(* IEC 61131-3 sources: model-first-plc-agent-ai/results/T2-W-22, 2 files *)

(* ---- a1_code.st ---- *)
FUNCTION_BLOCK FillingRuntime
VAR_INPUT
    start : BOOL;
    stop : BOOL;
    LSH : BOOL;
    LSHH : BOOL;
    TimerDuration : TIME;
END_VAR
VAR_OUTPUT
    fill_valve : BOOL;
    discharge_valve : BOOL;
END_VAR
VAR
    x0 : BOOL := TRUE;
    x1 : BOOL := FALSE;
    timer_done : BOOL := FALSE;
    FillingTimer : TON;
END_VAR

(* Admit a start event only from the initial situation. *)
IF x0 AND start AND NOT stop AND NOT LSHH THEN
    x0 := FALSE;
    x1 := TRUE;
END_IF;

(* Timing begins in the same scan that x1 becomes active. *)
FillingTimer(IN := x1, PT := TimerDuration);
timer_done := FillingTimer.Q;

(* Terminate filling before updating the physical output commands. *)
IF x1 AND (stop OR LSHH OR timer_done) THEN
    x1 := FALSE;
    x0 := TRUE;

    (* Reset immediately so a subsequent start receives a fresh interval. *)
    FillingTimer(IN := FALSE, PT := TimerDuration);
    timer_done := FALSE;
END_IF;

fill_valve := x1;
discharge_valve := FALSE;

END_FUNCTION_BLOCK

PROGRAM Main
VAR
    StartCommand AT %IX100.0 : BOOL;
    StopCommand AT %IX100.1 : BOOL;
    LSH AT %IX100.2 : BOOL;
    LSHH AT %IX100.3 : BOOL;
    FillValve AT %QX100.0 : BOOL;
    DischargeValve AT %QX100.1 : BOOL;
END_VAR
VAR
    (* Configurable filling interval. *)
    TimerDuration : TIME := T#5s;
    StartEdge : R_TRIG;
    FillingControl : FillingRuntime;
END_VAR

StartEdge(CLK := StartCommand);

FillingControl(
    start := StartEdge.Q,
    stop := StopCommand,
    LSH := LSH,
    LSHH := LSHH,
    TimerDuration := TimerDuration
);

FillValve := FillingControl.fill_valve;
DischargeValve := FillingControl.discharge_valve;

END_PROGRAM

(* ---- a2_code.st ---- *)
FUNCTION_BLOCK FB_TimedTank
VAR_INPUT
    StartCommand : BOOL;
    StopCommand : BOOL;
    LSH : BOOL;
    LSHH : BOOL;
    TimerDuration : TIME;
END_VAR
VAR_OUTPUT
    fill_valve : BOOL;
    discharge_valve : BOOL;
END_VAR
VAR
    StartEdge : R_TRIG;
    FillingTimer : TON;
    CycleState : INT := 0;
    start : BOOL;
    stop : BOOL;
    timer_done : BOOL;
END_VAR

StartEdge(CLK := StartCommand);
start := StartEdge.Q;
stop := StopCommand;

IF stop THEN
    CycleState := 0;
ELSE
    CASE CycleState OF
        0:
            IF start AND NOT LSHH THEN
                CycleState := 1;
            END_IF;
        1:
            IF LSHH THEN
                CycleState := 0;
            END_IF;
    ELSE
        CycleState := 0;
    END_CASE;
END_IF;

(* Start timing in the same scan that the filling step becomes active. *)
FillingTimer(IN := (CycleState = 1), PT := TimerDuration);
timer_done := FillingTimer.Q;

IF (CycleState = 1) AND timer_done THEN
    CycleState := 0;

    (* Reset the owned timer immediately upon leaving the filling step. *)
    FillingTimer(IN := FALSE, PT := TimerDuration);
    timer_done := FillingTimer.Q;
END_IF;

fill_valve := (CycleState = 1);
discharge_valve := FALSE;

END_FUNCTION_BLOCK

PROGRAM Main
VAR
    StartCommand AT %IX100.0 : BOOL;
    StopCommand AT %IX100.1 : BOOL;
    LSH AT %IX100.2 : BOOL;
    LSHH AT %IX100.3 : BOOL;
    FillValve AT %QX100.0 : BOOL;
    DischargeValve AT %QX100.1 : BOOL;
END_VAR
VAR
    TankController : FB_TimedTank;
    TimerDuration : TIME := T#5s;
END_VAR

TankController(
    StartCommand := StartCommand,
    StopCommand := StopCommand,
    LSH := LSH,
    LSHH := LSHH,
    TimerDuration := TimerDuration
);

FillValve := TankController.fill_valve;
DischargeValve := TankController.discharge_valve;

END_PROGRAM
